FUNCTION_BLOCK AirLockCmd (* Emergencia: abre a AV-4x171 (air fill) no inicio da aeracao durante o AirLockTime *)
  (* Standard: 61499-2 *)
  (* Version 1.1, 30/10/2026, Hidryco, Hidryco, 1.1: so em Mode 3; o tempo conta da confirmacao de aberta da AV-4x171 (FB_VALVE/Opened) e nao mais do Starting; fecha no fim do tempo, quando a fase sai ou quando o modo sai de 3; sem o reenvio no Run (o seletor so repassa mudancas). 1.0: pulso AirLock no inicio da fase de aeracao durante AirLockTime. AirLockTime = 0 nao abre. *)
  PACKAGE SE.Nereda;
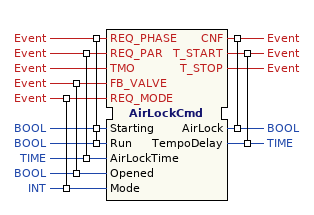
  EVENT_INPUT
    REQ_PHASE WITH Starting, Run; (* Estado da fase de aeracao (IPhase.Interlocked_CNF) *)
    REQ_PAR WITH AirLockTime; (* Tempo de air lock da emergencia *)
    TMO; (* Fim do tempo (E_DELAY.EO) *)
    FB_VALVE WITH Opened; (* Retorno da AV-4x171 *)
    REQ_MODE WITH Mode; (* Modo da planta *)
  END_EVENT
  EVENT_OUTPUT
    CNF WITH AirLock; (* AirLock mudou *)
    T_START WITH TempoDelay; (* Inicia o E_DELAY *)
    T_STOP; (* Para o E_DELAY *)
  END_EVENT
  VAR_INPUT
    Starting : BOOL; (* Fase de aeracao partindo *)
    Run : BOOL; (* Fase de aeracao rodando *)
    AirLockTime : TIME; (* Tempo de abertura da AV-4x171 no inicio da aeracao (emergencia) *)
    Opened : BOOL; (* AV-4x171 aberta *)
    Mode : INT; (* Modo da planta (3 = emergencia) *)
  END_VAR
  VAR_OUTPUT
    AirLock : BOOL; (* TRUE = AV-4x171 aberta pelo air lock *)
    TempoDelay : TIME; (* Tempo para o E_DELAY *)
  END_VAR
  VAR
    bAtivo : BOOL; (* Fase ativa na ultima leitura *)
    bAbrir : BOOL;
    bFechar : BOOL;
    bContando : BOOL; (* E_DELAY do AirLockTime em andamento (valvula ja confirmou aberta) *)
  END_VAR
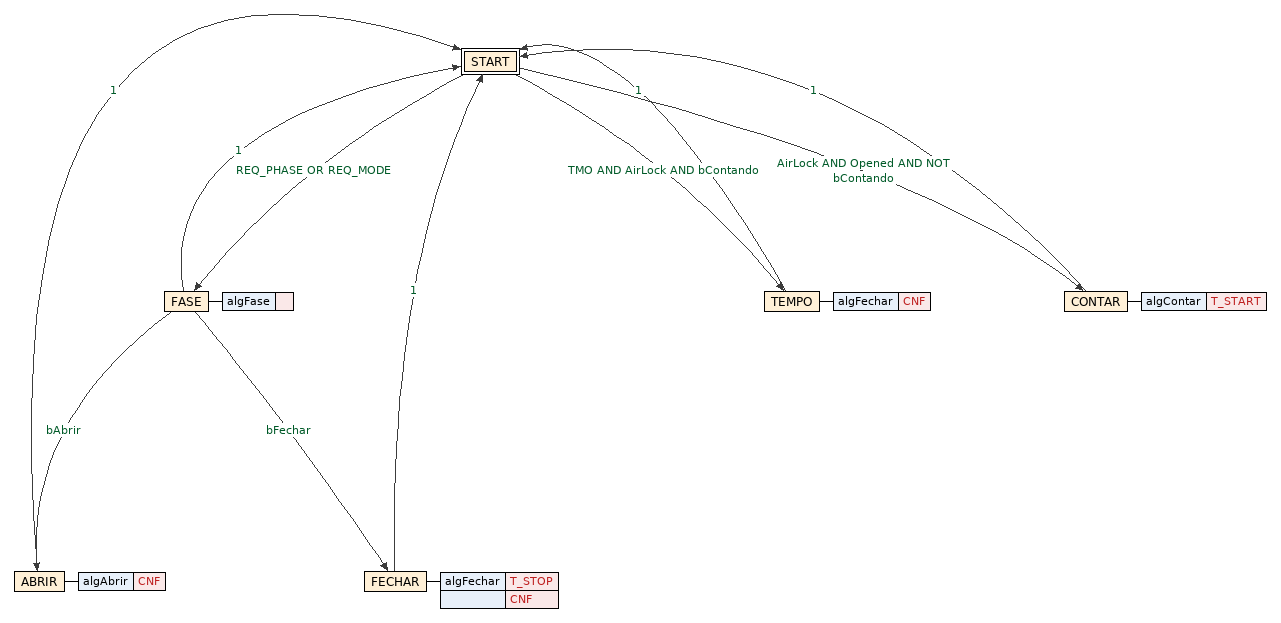
  EC_STATES
    START; (* Initial State *)
    FASE : algFase;
    ABRIR : algAbrir -> CNF;
    FECHAR : algFechar -> T_STOP, -> CNF;
    CONTAR : algContar -> T_START; (* Valvula aberta: inicia o AirLockTime *)
    TEMPO : algFechar -> CNF;
  END_STATES
  EC_TRANSITIONS
    START TO FASE := REQ_PHASE OR REQ_MODE;
    FASE TO ABRIR := bAbrir;
    FASE TO FECHAR := bFechar;
    FASE TO START := 1;
    ABRIR TO START := 1;
    FECHAR TO START := 1;
    START TO TEMPO := TMO AND AirLock AND bContando;
    TEMPO TO START := 1;
    START TO CONTAR := AirLock AND Opened AND NOT bContando;
    CONTAR TO START := 1;
  END_TRANSITIONS
  ALGORITHM algFase IN ST:
(* Abre no flanco de subida da fase (Starting ou Run), so em Mode 3 e se houver tempo;
   fecha quando a fase sai ou o modo sai de 3 *)
bAbrir := (Starting OR Run) AND NOT bAtivo AND (AirLockTime > T#0ms) AND (Mode = 3) AND NOT AirLock;
bFechar := (NOT (Starting OR Run) OR (Mode <> 3)) AND AirLock;
bAtivo := Starting OR Run;
  END_ALGORITHM
  ALGORITHM algAbrir IN ST:
AirLock := TRUE;
bContando := FALSE;
  END_ALGORITHM
  ALGORITHM algFechar IN ST:
AirLock := FALSE;
bContando := FALSE;
  END_ALGORITHM
  ALGORITHM algContar IN ST:
bContando := TRUE;
TempoDelay := AirLockTime;
  END_ALGORITHM
END_FUNCTION_BLOCK
